// TIA Portal V15.1 export
FUNCTION "Common" : Void   // FC1, LAD
TITLE = Common
{ S7_Optimized_Access := 'TRUE' }
VERSION : 0.1
// E-STOP latch, RESET edge, parameter check (decisions/0006)
// stored: AutoNumber false, IsIECCheckEnabled false, SetENOAutomatically False
   VAR_TEMP   // added for the SCL form of the ladder/FBD networks
      _w1 : Bool;
   END_VAR
BEGIN

REGION Network 1: R-06 — RESET edge (not on first scan)
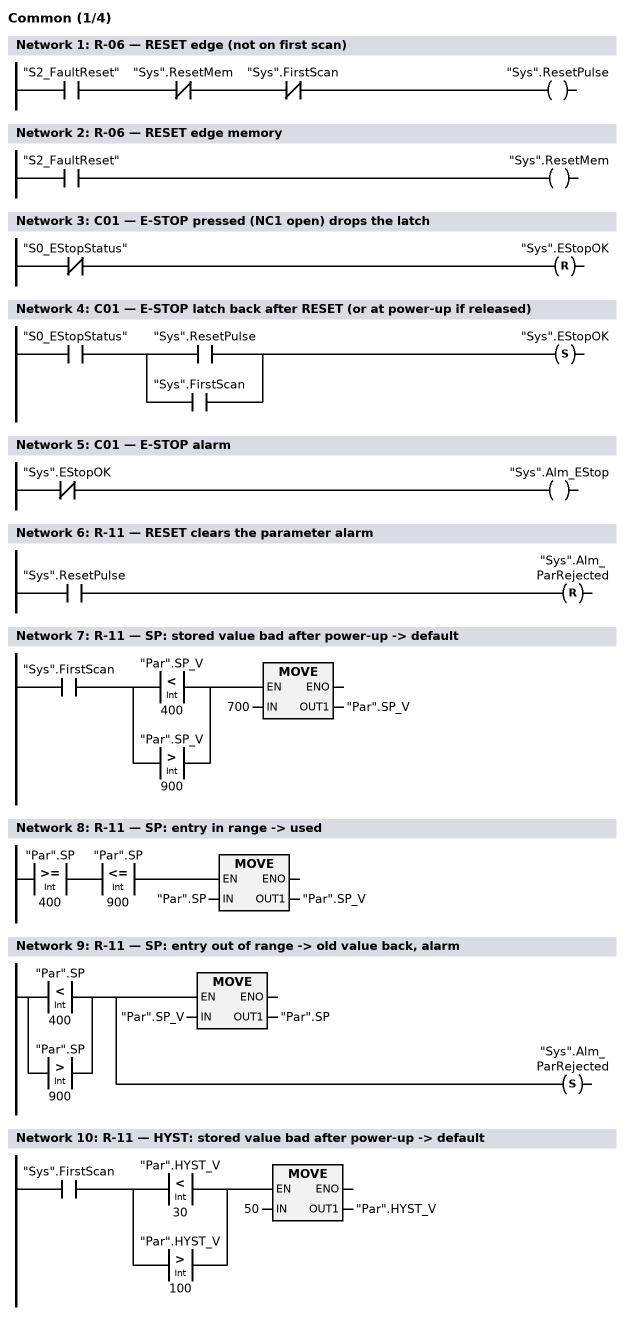
   RUNG wire#powerrail
      Contact( "S2_FaultReset" )
      I_Contact( "Sys".ResetMem )
      I_Contact( "Sys".FirstScan )
      Coil( "Sys".ResetPulse )
   END_RUNG
   // the same network as SCL:
   "Sys".ResetPulse := "S2_FaultReset" AND NOT "Sys".ResetMem AND NOT "Sys".FirstScan;
END_REGION

REGION Network 2: R-06 — RESET edge memory
   RUNG wire#powerrail
      Contact( "S2_FaultReset" )
      Coil( "Sys".ResetMem )
   END_RUNG
   // the same network as SCL:
   "Sys".ResetMem := "S2_FaultReset";
END_REGION

REGION Network 3: C01 — E-STOP pressed (NC1 open) drops the latch
   RUNG wire#powerrail
      I_Contact( "S0_EStopStatus" )
      R_Coil( "Sys".EStopOK )
   END_RUNG
   // the same network as SCL:
   IF NOT "S0_EStopStatus" THEN "Sys".EStopOK := FALSE; END_IF;
END_REGION

REGION Network 4: C01 — E-STOP latch back after RESET (or at power-up if released)
   RUNG wire#powerrail
      Contact( "S0_EStopStatus" )
      wire#w1
      Contact( "Sys".ResetPulse )
      wire#w2
      S_Coil( "Sys".EStopOK )
   END_RUNG
   RUNG wire#w1
      Contact( "Sys".FirstScan )
   END_RUNG wire#w2
   // the same network as SCL:
   IF "S0_EStopStatus" AND ("Sys".ResetPulse OR "Sys".FirstScan) THEN "Sys".EStopOK := TRUE; END_IF;
END_REGION

REGION Network 5: C01 — E-STOP alarm
   RUNG wire#powerrail
      I_Contact( "Sys".EStopOK )
      Coil( "Sys".Alm_EStop )
   END_RUNG
   // the same network as SCL:
   "Sys".Alm_EStop := NOT "Sys".EStopOK;
END_REGION

REGION Network 6: R-11 — RESET clears the parameter alarm
   RUNG wire#powerrail
      Contact( "Sys".ResetPulse )
      R_Coil( "Sys".Alm_ParRejected )
   END_RUNG
   // the same network as SCL:
   IF "Sys".ResetPulse THEN "Sys".Alm_ParRejected := FALSE; END_IF;
END_REGION

REGION Network 7: R-11 — SP: stored value bad after power-up -> default
   RUNG wire#powerrail
      Contact( "Sys".FirstScan )
      wire#w1
      { S7_Templates := "SrcType := Int" } LT_Contact(in1 := "Par".SP_V, in2 := 400)
      wire#w2
      { S7_GenerateENO := "TRUE" } Move(in := 700, out1 => "Par".SP_V)
   END_RUNG
   RUNG wire#w1
      { S7_Templates := "SrcType := Int" } GT_Contact(in1 := "Par".SP_V, in2 := 900)
   END_RUNG wire#w2
   // the same network as SCL:
   IF "Sys".FirstScan AND (("Par".SP_V < 400) OR ("Par".SP_V > 900)) THEN "Par".SP_V := 700; END_IF;
END_REGION

REGION Network 8: R-11 — SP: entry in range -> used
   RUNG wire#powerrail
      { S7_Templates := "SrcType := Int" } GE_Contact(in1 := "Par".SP, in2 := 400)
      { S7_Templates := "SrcType := Int" } LE_Contact(in1 := "Par".SP, in2 := 900)
      { S7_GenerateENO := "TRUE" } Move(in := "Par".SP, out1 => "Par".SP_V)
   END_RUNG
   // the same network as SCL:
   IF ("Par".SP >= 400) AND ("Par".SP <= 900) THEN "Par".SP_V := "Par".SP; END_IF;
END_REGION

REGION Network 9: R-11 — SP: entry out of range -> old value back, alarm
   RUNG wire#powerrail
      { S7_Templates := "SrcType := Int" } LT_Contact(in1 := "Par".SP, in2 := 400)
      wire#w1
      { S7_GenerateENO := "TRUE" } Move(in := "Par".SP_V, out1 => "Par".SP)
   END_RUNG
   RUNG wire#powerrail
      { S7_Templates := "SrcType := Int" } GT_Contact(in1 := "Par".SP, in2 := 900)
   END_RUNG wire#w1
   RUNG wire#w1
      S_Coil( "Sys".Alm_ParRejected )
   END_RUNG
   // the same network as SCL:
   #_w1 := ("Par".SP < 400) OR ("Par".SP > 900);
   IF #_w1 THEN
       "Par".SP := "Par".SP_V;
       "Sys".Alm_ParRejected := TRUE;
   END_IF;
END_REGION

REGION Network 10: R-11 — HYST: stored value bad after power-up -> default
   RUNG wire#powerrail
      Contact( "Sys".FirstScan )
      wire#w1
      { S7_Templates := "SrcType := Int" } LT_Contact(in1 := "Par".HYST_V, in2 := 30)
      wire#w2
      { S7_GenerateENO := "TRUE" } Move(in := 50, out1 => "Par".HYST_V)
   END_RUNG
   RUNG wire#w1
      { S7_Templates := "SrcType := Int" } GT_Contact(in1 := "Par".HYST_V, in2 := 100)
   END_RUNG wire#w2
   // the same network as SCL:
   IF "Sys".FirstScan AND (("Par".HYST_V < 30) OR ("Par".HYST_V > 100)) THEN "Par".HYST_V := 50; END_IF;
END_REGION

REGION Network 11: R-11 — HYST: entry in range -> used
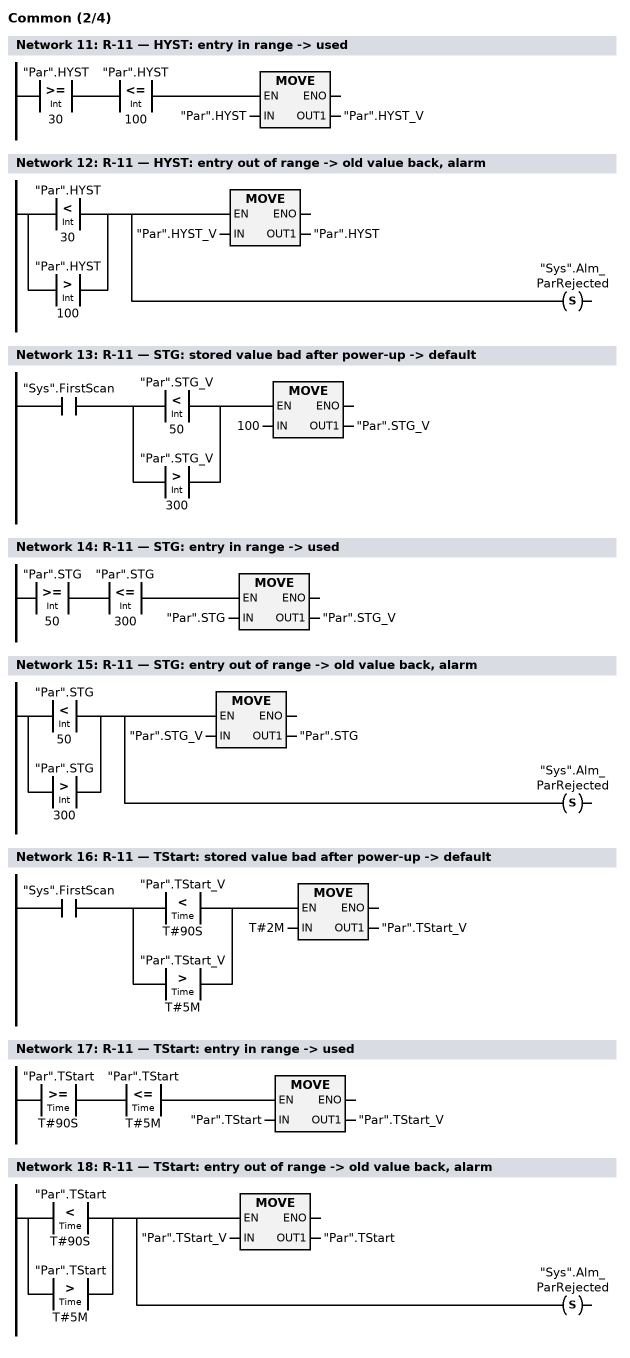
   RUNG wire#powerrail
      { S7_Templates := "SrcType := Int" } GE_Contact(in1 := "Par".HYST, in2 := 30)
      { S7_Templates := "SrcType := Int" } LE_Contact(in1 := "Par".HYST, in2 := 100)
      { S7_GenerateENO := "TRUE" } Move(in := "Par".HYST, out1 => "Par".HYST_V)
   END_RUNG
   // the same network as SCL:
   IF ("Par".HYST >= 30) AND ("Par".HYST <= 100) THEN "Par".HYST_V := "Par".HYST; END_IF;
END_REGION

REGION Network 12: R-11 — HYST: entry out of range -> old value back, alarm
   RUNG wire#powerrail
      { S7_Templates := "SrcType := Int" } LT_Contact(in1 := "Par".HYST, in2 := 30)
      wire#w1
      { S7_GenerateENO := "TRUE" } Move(in := "Par".HYST_V, out1 => "Par".HYST)
   END_RUNG
   RUNG wire#powerrail
      { S7_Templates := "SrcType := Int" } GT_Contact(in1 := "Par".HYST, in2 := 100)
   END_RUNG wire#w1
   RUNG wire#w1
      S_Coil( "Sys".Alm_ParRejected )
   END_RUNG
   // the same network as SCL:
   #_w1 := ("Par".HYST < 30) OR ("Par".HYST > 100);
   IF #_w1 THEN
       "Par".HYST := "Par".HYST_V;
       "Sys".Alm_ParRejected := TRUE;
   END_IF;
END_REGION

REGION Network 13: R-11 — STG: stored value bad after power-up -> default
   RUNG wire#powerrail
      Contact( "Sys".FirstScan )
      wire#w1
      { S7_Templates := "SrcType := Int" } LT_Contact(in1 := "Par".STG_V, in2 := 50)
      wire#w2
      { S7_GenerateENO := "TRUE" } Move(in := 100, out1 => "Par".STG_V)
   END_RUNG
   RUNG wire#w1
      { S7_Templates := "SrcType := Int" } GT_Contact(in1 := "Par".STG_V, in2 := 300)
   END_RUNG wire#w2
   // the same network as SCL:
   IF "Sys".FirstScan AND (("Par".STG_V < 50) OR ("Par".STG_V > 300)) THEN "Par".STG_V := 100; END_IF;
END_REGION

REGION Network 14: R-11 — STG: entry in range -> used
   RUNG wire#powerrail
      { S7_Templates := "SrcType := Int" } GE_Contact(in1 := "Par".STG, in2 := 50)
      { S7_Templates := "SrcType := Int" } LE_Contact(in1 := "Par".STG, in2 := 300)
      { S7_GenerateENO := "TRUE" } Move(in := "Par".STG, out1 => "Par".STG_V)
   END_RUNG
   // the same network as SCL:
   IF ("Par".STG >= 50) AND ("Par".STG <= 300) THEN "Par".STG_V := "Par".STG; END_IF;
END_REGION

REGION Network 15: R-11 — STG: entry out of range -> old value back, alarm
   RUNG wire#powerrail
      { S7_Templates := "SrcType := Int" } LT_Contact(in1 := "Par".STG, in2 := 50)
      wire#w1
      { S7_GenerateENO := "TRUE" } Move(in := "Par".STG_V, out1 => "Par".STG)
   END_RUNG
   RUNG wire#powerrail
      { S7_Templates := "SrcType := Int" } GT_Contact(in1 := "Par".STG, in2 := 300)
   END_RUNG wire#w1
   RUNG wire#w1
      S_Coil( "Sys".Alm_ParRejected )
   END_RUNG
   // the same network as SCL:
   #_w1 := ("Par".STG < 50) OR ("Par".STG > 300);
   IF #_w1 THEN
       "Par".STG := "Par".STG_V;
       "Sys".Alm_ParRejected := TRUE;
   END_IF;
END_REGION

REGION Network 16: R-11 — TStart: stored value bad after power-up -> default
   RUNG wire#powerrail
      Contact( "Sys".FirstScan )
      wire#w1
      { S7_Templates := "SrcType := Time" } LT_Contact(in1 := "Par".TStart_V, in2 := T#90S)
      wire#w2
      { S7_GenerateENO := "TRUE" } Move(in := T#2M, out1 => "Par".TStart_V)
   END_RUNG
   RUNG wire#w1
      { S7_Templates := "SrcType := Time" } GT_Contact(in1 := "Par".TStart_V, in2 := T#5M)
   END_RUNG wire#w2
   // the same network as SCL:
   IF "Sys".FirstScan AND (("Par".TStart_V < T#90S) OR ("Par".TStart_V > T#5M)) THEN
       "Par".TStart_V := T#2M;
   END_IF;
END_REGION

REGION Network 17: R-11 — TStart: entry in range -> used
   RUNG wire#powerrail
      { S7_Templates := "SrcType := Time" } GE_Contact(in1 := "Par".TStart, in2 := T#90S)
      { S7_Templates := "SrcType := Time" } LE_Contact(in1 := "Par".TStart, in2 := T#5M)
      { S7_GenerateENO := "TRUE" } Move(in := "Par".TStart, out1 => "Par".TStart_V)
   END_RUNG
   // the same network as SCL:
   IF ("Par".TStart >= T#90S) AND ("Par".TStart <= T#5M) THEN "Par".TStart_V := "Par".TStart; END_IF;
END_REGION

REGION Network 18: R-11 — TStart: entry out of range -> old value back, alarm
   RUNG wire#powerrail
      { S7_Templates := "SrcType := Time" } LT_Contact(in1 := "Par".TStart, in2 := T#90S)
      wire#w1
      { S7_GenerateENO := "TRUE" } Move(in := "Par".TStart_V, out1 => "Par".TStart)
   END_RUNG
   RUNG wire#powerrail
      { S7_Templates := "SrcType := Time" } GT_Contact(in1 := "Par".TStart, in2 := T#5M)
   END_RUNG wire#w1
   RUNG wire#w1
      S_Coil( "Sys".Alm_ParRejected )
   END_RUNG
   // the same network as SCL:
   #_w1 := ("Par".TStart < T#90S) OR ("Par".TStart > T#5M);
   IF #_w1 THEN
       "Par".TStart := "Par".TStart_V;
       "Sys".Alm_ParRejected := TRUE;
   END_IF;
END_REGION

REGION Network 19: R-11 — TDrnOn: stored value bad after power-up -> default
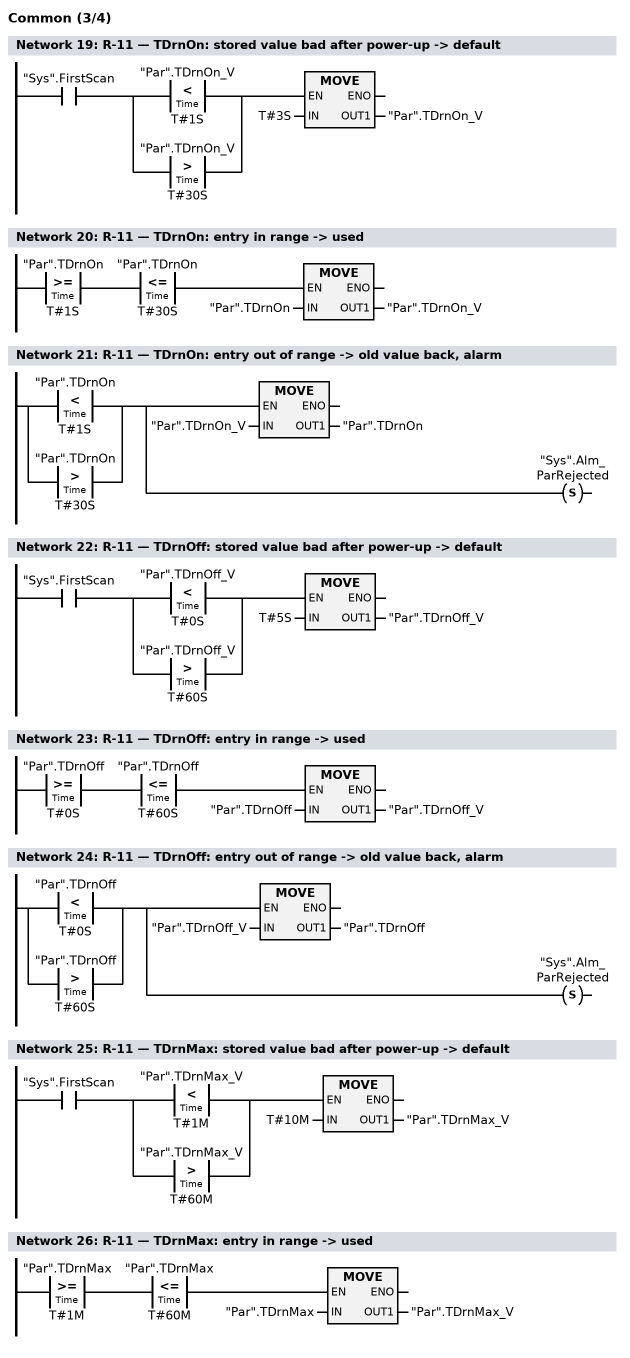
   RUNG wire#powerrail
      Contact( "Sys".FirstScan )
      wire#w1
      { S7_Templates := "SrcType := Time" } LT_Contact(in1 := "Par".TDrnOn_V, in2 := T#1S)
      wire#w2
      { S7_GenerateENO := "TRUE" } Move(in := T#3S, out1 => "Par".TDrnOn_V)
   END_RUNG
   RUNG wire#w1
      { S7_Templates := "SrcType := Time" } GT_Contact(in1 := "Par".TDrnOn_V, in2 := T#30S)
   END_RUNG wire#w2
   // the same network as SCL:
   IF "Sys".FirstScan AND (("Par".TDrnOn_V < T#1S) OR ("Par".TDrnOn_V > T#30S)) THEN
       "Par".TDrnOn_V := T#3S;
   END_IF;
END_REGION

REGION Network 20: R-11 — TDrnOn: entry in range -> used
   RUNG wire#powerrail
      { S7_Templates := "SrcType := Time" } GE_Contact(in1 := "Par".TDrnOn, in2 := T#1S)
      { S7_Templates := "SrcType := Time" } LE_Contact(in1 := "Par".TDrnOn, in2 := T#30S)
      { S7_GenerateENO := "TRUE" } Move(in := "Par".TDrnOn, out1 => "Par".TDrnOn_V)
   END_RUNG
   // the same network as SCL:
   IF ("Par".TDrnOn >= T#1S) AND ("Par".TDrnOn <= T#30S) THEN "Par".TDrnOn_V := "Par".TDrnOn; END_IF;
END_REGION

REGION Network 21: R-11 — TDrnOn: entry out of range -> old value back, alarm
   RUNG wire#powerrail
      { S7_Templates := "SrcType := Time" } LT_Contact(in1 := "Par".TDrnOn, in2 := T#1S)
      wire#w1
      { S7_GenerateENO := "TRUE" } Move(in := "Par".TDrnOn_V, out1 => "Par".TDrnOn)
   END_RUNG
   RUNG wire#powerrail
      { S7_Templates := "SrcType := Time" } GT_Contact(in1 := "Par".TDrnOn, in2 := T#30S)
   END_RUNG wire#w1
   RUNG wire#w1
      S_Coil( "Sys".Alm_ParRejected )
   END_RUNG
   // the same network as SCL:
   #_w1 := ("Par".TDrnOn < T#1S) OR ("Par".TDrnOn > T#30S);
   IF #_w1 THEN
       "Par".TDrnOn := "Par".TDrnOn_V;
       "Sys".Alm_ParRejected := TRUE;
   END_IF;
END_REGION

REGION Network 22: R-11 — TDrnOff: stored value bad after power-up -> default
   RUNG wire#powerrail
      Contact( "Sys".FirstScan )
      wire#w1
      { S7_Templates := "SrcType := Time" } LT_Contact(in1 := "Par".TDrnOff_V, in2 := T#0S)
      wire#w2
      { S7_GenerateENO := "TRUE" } Move(in := T#5S, out1 => "Par".TDrnOff_V)
   END_RUNG
   RUNG wire#w1
      { S7_Templates := "SrcType := Time" } GT_Contact(in1 := "Par".TDrnOff_V, in2 := T#60S)
   END_RUNG wire#w2
   // the same network as SCL:
   IF "Sys".FirstScan AND (("Par".TDrnOff_V < T#0S) OR ("Par".TDrnOff_V > T#60S)) THEN
       "Par".TDrnOff_V := T#5S;
   END_IF;
END_REGION

REGION Network 23: R-11 — TDrnOff: entry in range -> used
   RUNG wire#powerrail
      { S7_Templates := "SrcType := Time" } GE_Contact(in1 := "Par".TDrnOff, in2 := T#0S)
      { S7_Templates := "SrcType := Time" } LE_Contact(in1 := "Par".TDrnOff, in2 := T#60S)
      { S7_GenerateENO := "TRUE" } Move(in := "Par".TDrnOff, out1 => "Par".TDrnOff_V)
   END_RUNG
   // the same network as SCL:
   IF ("Par".TDrnOff >= T#0S) AND ("Par".TDrnOff <= T#60S) THEN "Par".TDrnOff_V := "Par".TDrnOff; END_IF;
END_REGION

REGION Network 24: R-11 — TDrnOff: entry out of range -> old value back, alarm
   RUNG wire#powerrail
      { S7_Templates := "SrcType := Time" } LT_Contact(in1 := "Par".TDrnOff, in2 := T#0S)
      wire#w1
      { S7_GenerateENO := "TRUE" } Move(in := "Par".TDrnOff_V, out1 => "Par".TDrnOff)
   END_RUNG
   RUNG wire#powerrail
      { S7_Templates := "SrcType := Time" } GT_Contact(in1 := "Par".TDrnOff, in2 := T#60S)
   END_RUNG wire#w1
   RUNG wire#w1
      S_Coil( "Sys".Alm_ParRejected )
   END_RUNG
   // the same network as SCL:
   #_w1 := ("Par".TDrnOff < T#0S) OR ("Par".TDrnOff > T#60S);
   IF #_w1 THEN
       "Par".TDrnOff := "Par".TDrnOff_V;
       "Sys".Alm_ParRejected := TRUE;
   END_IF;
END_REGION

REGION Network 25: R-11 — TDrnMax: stored value bad after power-up -> default
   RUNG wire#powerrail
      Contact( "Sys".FirstScan )
      wire#w1
      { S7_Templates := "SrcType := Time" } LT_Contact(in1 := "Par".TDrnMax_V, in2 := T#1M)
      wire#w2
      { S7_GenerateENO := "TRUE" } Move(in := T#10M, out1 => "Par".TDrnMax_V)
   END_RUNG
   RUNG wire#w1
      { S7_Templates := "SrcType := Time" } GT_Contact(in1 := "Par".TDrnMax_V, in2 := T#60M)
   END_RUNG wire#w2
   // the same network as SCL:
   IF "Sys".FirstScan AND (("Par".TDrnMax_V < T#1M) OR ("Par".TDrnMax_V > T#60M)) THEN
       "Par".TDrnMax_V := T#10M;
   END_IF;
END_REGION

REGION Network 26: R-11 — TDrnMax: entry in range -> used
   RUNG wire#powerrail
      { S7_Templates := "SrcType := Time" } GE_Contact(in1 := "Par".TDrnMax, in2 := T#1M)
      { S7_Templates := "SrcType := Time" } LE_Contact(in1 := "Par".TDrnMax, in2 := T#60M)
      { S7_GenerateENO := "TRUE" } Move(in := "Par".TDrnMax, out1 => "Par".TDrnMax_V)
   END_RUNG
   // the same network as SCL:
   IF ("Par".TDrnMax >= T#1M) AND ("Par".TDrnMax <= T#60M) THEN "Par".TDrnMax_V := "Par".TDrnMax; END_IF;
END_REGION

REGION Network 27: R-11 — TDrnMax: entry out of range -> old value back, alarm
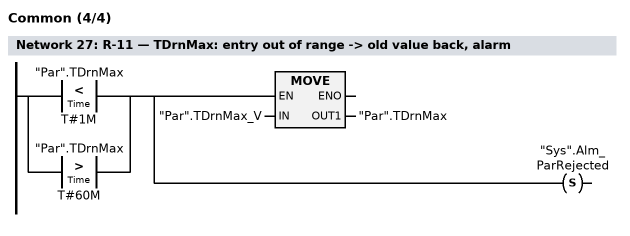
   RUNG wire#powerrail
      { S7_Templates := "SrcType := Time" } LT_Contact(in1 := "Par".TDrnMax, in2 := T#1M)
      wire#w1
      { S7_GenerateENO := "TRUE" } Move(in := "Par".TDrnMax_V, out1 => "Par".TDrnMax)
   END_RUNG
   RUNG wire#powerrail
      { S7_Templates := "SrcType := Time" } GT_Contact(in1 := "Par".TDrnMax, in2 := T#60M)
   END_RUNG wire#w1
   RUNG wire#w1
      S_Coil( "Sys".Alm_ParRejected )
   END_RUNG
   // the same network as SCL:
   #_w1 := ("Par".TDrnMax < T#1M) OR ("Par".TDrnMax > T#60M);
   IF #_w1 THEN
       "Par".TDrnMax := "Par".TDrnMax_V;
       "Sys".Alm_ParRejected := TRUE;
   END_IF;
END_REGION
END_FUNCTION
